SYSTEM test
  (* Standard: ISO 11783 / IEC 61499; ApplicationDomain: Slurry Tanker; Description: https://github.com/Meisterschulen-am-Ostbahnhof-Munchen/4diac-SlurryTanker-sample *)
  (* Version 0.1, 2022-11-10, Franz Höpfinger, Meisterschulen am Ostbahnhof, München, erste Version. *)
  (* Version 0.2, 2022-11-11, Franz Höpfinger, Meisterschulen am Ostbahnhof, München, Vorgewendeautomatik *)
  (* Version 0.3, 2022-11-16, Franz Höpfinger, Meisterschulen am Ostbahnhof, München, alle Zeiten auf T#3s *)
  DEVICE FORTE_PC : FORTE_PC(MGR_ID := C_00)
    {SET_ATTRIBUTE(Profile, HOLOBLOC)}
    {SET_ATTRIBUTE(FBType, E_SWITCH, E_SR_RETRIG, E_R_TRIG, E_T_FF, E_IMPULSE, E_SR, E_F_TRIG, E_REND, E_D_FF)} (* created during deployment *)
    RESOURCE EMB_RES : EMB_RES
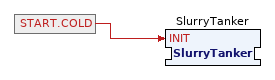
      SUBAPPS
        SlurryTanker : SlurryTanker;
      END_SUBAPPS
      EVENT_CONNECTIONS
        START.COLD TO SlurryTanker.INIT;
      END_CONNECTIONS
    END_RESOURCE
  END_DEVICE
  SEGMENTS
    Ethernet : Ethernet;
  END_SEGMENTS
  LINKS
    FORTE_PC => Ethernet;
  END_LINKS
END_SYSTEM
